// Tout ce qui porte un override et un état : machine, station, module, objet (docs/04 § 4)
INTERFACE I_Node

PROPERTY EffectiveOverride : LREAL
GET
END_GET
END_PROPERTY

PROPERTY NodeState : E_ObjState
GET
END_GET
END_PROPERTY

END_INTERFACE

(* stored: Version 1.1.0.1, ProductVersion 3.1.4024.12
   Itf I_Node: Id {09953dc9-61db-5736-8df7-50e1208b101f}
   Property EffectiveOverride: Id {bcef9c2e-644c-5bd3-8441-c2ab25811f90}
   Get Get: Id {84d9ca1b-1768-55b3-a0e2-e0f9424773d6}
   Property NodeState: Id {2e6d95bd-b3e1-5374-abb6-3606bce7fca0}
   Get Get: Id {b5674053-6f8b-5782-b00c-563ce7bb615c} *)
